# B&R Automation Studio project BasdfasdfKVBO0823_1
Automation Studio 4.5.2.102

## Configuration Config1

CPU 4PP065.0351-P74, AutomationRuntime D4.52, Build 4.1.2, Vc V4.52.0

### Task classes (Cpu.sw)
```
Cyclic#3:
  Program <- Program.prg
Binaries: udbdef, TCData, ashwd, User, asfw, arconfig, sysconf, Role, ashwac, iomap
Libraries: Library
```

### Hardware
```
4PP065_0351_P74 : 4PP065.0351-P74 v1.0.4.0
  Connector IF5:
    ActivateDevice = 1
    Mode = Manual
    InternetAddress = 10.0.1.10
    SubnetMask = 255.255.255.0
  ConfigurationID = labBR
  Simulation = 1
  KeyMappingFile = VC\4PP065_0351_P74.dis
```

- Physical/Config1/4PP065_0351_P74/IoMap.iom: same as Physical/Config1/4PP065_0351_P74/Cpu.per
- Physical/Config1/4PP065_0351_P74/PvMap.vvm: same as Physical/Config1/4PP065_0351_P74/Cpu.per
## Logical view

Binary libraries used (declarations not repeated): operator, runtime, astime, AsIecCon


### Program Logical/Program (ANSIC)

#### Cyclic.c - Cyclic code
```c
#include <bur/plctypes.h>

#ifdef _DEFAULT_INCLUDES
#include <AsDefault.h>
#endif

void _CYCLIC ProgramCyclic(void)
{
	REAL PI = 3.141592653589793;
	REAL desired_w = speed * 2.0 * PI / 60.0;
	speed_in_rad = desired_w;

	if (enable == 1){
		counter += 1;
		if ((counter >= 500 ) && (counter <= 1000)) speed = 70;
		else speed = 0;
	}
	else speed = 0;

	fb_controller.e = desired_w - fb_motor.w;
	FB_Regulator(&fb_controller);
	fb_motor.u = fb_controller.u;

	fb_motor_2.u = desired_w * fb_motor_2.ke;

	FB_Motor(&fb_motor);
	FB_Motor(&fb_motor_2);

}
```

#### Init.c - Initialization code
```c
#include <bur/plctypes.h>

#ifdef _DEFAULT_INCLUDES
#include <AsDefault.h>
#endif

void _INIT ProgramInit(void)
{
	enable = 1;
	counter = 0;
	speed = 0;
	speed_in_rad = 0;

	fb_motor.dt=0.002;
	fb_motor.ke=0.00096;
	fb_motor.Tm=0.04;
	fb_motor.integrator.dt = 0.002;
	fb_motor.sensor.dt = 0.002;

	fb_motor_2.dt = 0.002;
	fb_motor_2.ke = 0.00096;
	fb_motor_2.Tm = 0.04;
	fb_motor_2.integrator.dt = 0.002;
	fb_motor_2.sensor.dt = 0.002;

	fb_controller.dt=0.002;
	fb_controller.k_p = 0.0064;
	fb_controller.k_i = 0.16;
	fb_controller.max_abs_value=24;
	fb_controller.integrator.dt = 0.002;
}
```

#### Exit.c - Exit code
```c
#include <bur/plctypes.h>

#ifdef _DEFAULT_INCLUDES
	#include <AsDefault.h>
#endif

void _EXIT ProgramExit(void)
{

}
```

#### Variables.var - Local variables
```iecst
VAR
	counter : UDINT;
	fb_controller : FB_Regulator;
	fb_motor : FB_Motor;
	speed : UINT;
	enable : USINT;
	speed_in_rad : REAL;
	fb_motor_2 : FB_Motor;
END_VAR
```

### Library Logical/Library (ANSIC)

#### Library.fun - Exported functions and function blocks
```iecst
{REDUND_OK} FUNCTION_BLOCK FB_Regulator (*TODO: Add your comment here*) (*$GROUP=User,$CAT=User,$GROUPICON=User.png,$CATICON=User.png*)
	VAR_INPUT
		e : REAL;
	END_VAR
	VAR_OUTPUT
		u : REAL;
	END_VAR
	VAR
		k_p : REAL;
		k_i : REAL;
		integrator : FB_Integrator;
		iyOld : REAL;
		max_abs_value : REAL;
		dt : REAL;
	END_VAR
END_FUNCTION_BLOCK

{REDUND_OK} FUNCTION_BLOCK FB_Motor (*TODO: Add your comment here*) (*$GROUP=User,$CAT=User,$GROUPICON=User.png,$CATICON=User.png*)
	VAR_INPUT
		u : REAL;
	END_VAR
	VAR_OUTPUT
		w : REAL;
		phi : REAL;
	END_VAR
	VAR
		integrator : FB_Integrator;
		Tm : REAL;
		ke : REAL;
		dt : REAL;
		sensor : FB_Integrator;
	END_VAR
END_FUNCTION_BLOCK

{REDUND_OK} FUNCTION_BLOCK FB_Integrator (*TODO: Add your comment here*) (*$GROUP=User,$CAT=User,$GROUPICON=User.png,$CATICON=User.png*)
	VAR_INPUT
		in : REAL;
	END_VAR
	VAR_OUTPUT
		out : REAL;
	END_VAR
	VAR
		dt : REAL;
	END_VAR
	VAR_OUTPUT
		state : REAL;
	END_VAR
END_FUNCTION_BLOCK
```

#### FB_Regulator.c
```c
#include <bur/plctypes.h>
#ifdef __cplusplus
	extern "C"
	{
#endif
#include "Library.h"
#ifdef __cplusplus
	};
#endif
/* REGULATOR */
void FB_Regulator(struct FB_Regulator* inst)
{
	REAL p_part = inst->e * inst->k_p;

	REAL i_part = inst->e * inst->k_i;

	inst->integrator.in = i_part;

	FB_Integrator(&inst->integrator);

	i_part = inst->integrator.out;

	REAL total_output = p_part + i_part;

	if (total_output > inst->max_abs_value)
	{
		inst->u = inst->max_abs_value;
		inst->integrator.out = inst->max_abs_value - p_part;

	} else if (total_output < -inst->max_abs_value)
	{
		inst->u = -inst->max_abs_value;
		inst->integrator.out = -inst->max_abs_value - p_part;
	} else
	{
		inst->u = total_output;

	}
	inst->iyOld = i_part;
}
```

#### FB_Motor.c
```c
#include <bur/plctypes.h>
#ifdef __cplusplus
	extern "C"
	{
#endif
#include "Library.h"
#ifdef __cplusplus
	};
#endif
/* MOTOR */
void FB_Motor(struct FB_Motor* inst)
{
	REAL b1 = inst->u * (1/inst->ke) - inst->w;
	REAL b2 = b1/ inst->Tm;

	inst->integrator.in = b2;
	FB_Integrator(&inst->integrator);

	inst->w = inst->integrator.out;

	inst->sensor.in = inst->w;
	FB_Integrator(&inst->sensor);

	inst->phi = inst->sensor.out ;

}
```

#### FB_Integrator.c
```c
#include <bur/plctypes.h>
#ifdef __cplusplus
	extern "C"
	{
#endif
#include "Library.h"
#ifdef __cplusplus
	};
#endif
/* INTEGRATOR */
void FB_Integrator(struct FB_Integrator* inst)
{
	inst->out = inst->dt * inst->in + inst->state;
	inst->state = inst->out;
}
```
